SUBAPPLICATION SubApp_PC_A (* Geraet A: Variablen per CLIENT (opcua.adoc): Input_I1 schreibt 42 auf Increment (CLIENT_1_0), liest danach Incremented = 43 (CLIENT_0_1) *)
  (* Standard: 61499-2; Description: Copyright (c) 2026 Meisterschulen am Ostbahnhof This program and the accompanying materials are made available under the terms of the Eclipse Public License 2.0 which is available at https://www.eclipse.org/legal/epl-2.0/ SPDX-License-Identifier: EPL-2.0 *)
  (* Version 1.0, 2026-10-18, Franz Höpfinger, Meisterschulen am Ostbahnhof, opcua.adoc-Beispiel auf zwei Geraeten *)
  PACKAGE subapp::Training_16_OPC_UA_RES;
  IMPORT VV::const::OPC_UA::myOpcUaAddresses::T16_INC_CLIENT_WRITE;
  IMPORT VV::const::OPC_UA::myOpcUaAddresses::T16_INCD_CLIENT_READ;
  IMPORT logiBUS::io::DI::logiBUS_DI::Input_I1;
  IMPORT logiBUS::io::DI::logiBUS_DI_Events::BUTTON_PRESS_DOWN;
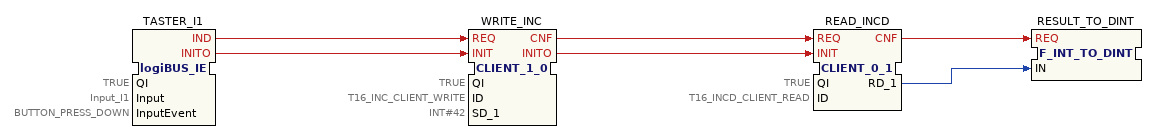
  FBS
    TASTER_I1 : logiBUS::io::DI::logiBUS_IE(QI := TRUE, Input := Input_I1, InputEvent := BUTTON_PRESS_DOWN);
    WRITE_INC : iec61499::net::CLIENT_1_0(QI := TRUE, ID := T16_INC_CLIENT_WRITE, SD_1 := INT#42);
    READ_INCD : iec61499::net::CLIENT_0_1(QI := TRUE, ID := T16_INCD_CLIENT_READ);
    RESULT_TO_DINT : iec61131::conversion::F_INT_TO_DINT;
  END_FBS
  EVENT_CONNECTIONS
    TASTER_I1.IND TO WRITE_INC.REQ;
    WRITE_INC.CNF TO READ_INCD.REQ;
    TASTER_I1.INITO TO WRITE_INC.INIT;
    WRITE_INC.INITO TO READ_INCD.INIT;
    READ_INCD.CNF TO RESULT_TO_DINT.REQ;
  END_CONNECTIONS
  DATA_CONNECTIONS
    READ_INCD.RD_1 TO RESULT_TO_DINT.IN;
  END_CONNECTIONS
END_SUBAPPLICATION
